(* IEC 61131-3 sources: rusty/tests/lit/single/type_promotion/bit_string/case_selector, 5 files *)

(* ---- byte_range_across_midpoint.st ---- *)
// RUN: %COMPILE %s && %RUN | %CHECK %s
// A range label that crosses the signed midpoint of the BYTE selector matches every value between its bounds.
FUNCTION branch : DINT
    VAR_INPUT
        x : BYTE;
    END_VAR

    CASE x OF
        16#00:
            branch := 1;
        16#01..16#09:
            branch := 2;
        16#0B..16#FE:
            branch := 3;
        16#FF:
            branch := 4;
    ELSE
        branch := 9;
    END_CASE
END_FUNCTION

FUNCTION main : DINT
    printf('16#00 -> %d$N', branch(16#00));                     // CHECK: 16#00 -> 1
    printf('16#05 -> %d$N', branch(16#05));                     // CHECK-NEXT: 16#05 -> 2
    printf('16#0A -> %d$N', branch(16#0A));                     // CHECK-NEXT: 16#0A -> 9
    printf('16#0B -> %d$N', branch(16#0B));                     // CHECK-NEXT: 16#0B -> 3
    printf('16#7F -> %d$N', branch(16#7F));                     // CHECK-NEXT: 16#7F -> 3
    printf('16#80 -> %d$N', branch(16#80));                     // CHECK-NEXT: 16#80 -> 3
    printf('16#C8 -> %d$N', branch(16#C8));                     // CHECK-NEXT: 16#C8 -> 3
    printf('16#FE -> %d$N', branch(16#FE));                     // CHECK-NEXT: 16#FE -> 3
    printf('16#FF -> %d$N', branch(16#FF));                     // CHECK-NEXT: 16#FF -> 4
END_FUNCTION

(* ---- dword_range_across_midpoint.st ---- *)
// RUN: %COMPILE %s && %RUN | %CHECK %s
// A range label that crosses the signed midpoint of the DWORD selector matches every value between its bounds.
FUNCTION branch : DINT
    VAR_INPUT
        x : DWORD;
    END_VAR

    CASE x OF
        16#0000_0000:
            branch := 1;
        16#0000_0001..16#0000_0009:
            branch := 2;
        16#0000_000B..16#FFFF_FFFE:
            branch := 3;
        16#FFFF_FFFF:
            branch := 4;
    ELSE
        branch := 9;
    END_CASE
END_FUNCTION

FUNCTION main : DINT
    printf('16#0000_0000 -> %d$N', branch(16#0000_0000));       // CHECK: 16#0000_0000 -> 1
    printf('16#0000_0005 -> %d$N', branch(16#0000_0005));       // CHECK-NEXT: 16#0000_0005 -> 2
    printf('16#0000_000A -> %d$N', branch(16#0000_000A));       // CHECK-NEXT: 16#0000_000A -> 9
    printf('16#0000_000B -> %d$N', branch(16#0000_000B));       // CHECK-NEXT: 16#0000_000B -> 3
    printf('16#7FFF_FFFF -> %d$N', branch(16#7FFF_FFFF));       // CHECK-NEXT: 16#7FFF_FFFF -> 3
    printf('16#8000_0000 -> %d$N', branch(16#8000_0000));       // CHECK-NEXT: 16#8000_0000 -> 3
    printf('16#B2D0_5E00 -> %d$N', branch(16#B2D0_5E00));       // CHECK-NEXT: 16#B2D0_5E00 -> 3
    printf('16#FFFF_FFFE -> %d$N', branch(16#FFFF_FFFE));       // CHECK-NEXT: 16#FFFF_FFFE -> 3
    printf('16#FFFF_FFFF -> %d$N', branch(16#FFFF_FFFF));       // CHECK-NEXT: 16#FFFF_FFFF -> 4
END_FUNCTION

(* ---- lword_range_across_midpoint.st ---- *)
// RUN: %COMPILE %s && %RUN | %CHECK %s
// A range label that crosses the signed midpoint of the LWORD selector matches every value between its bounds.
FUNCTION branch : DINT
    VAR_INPUT
        x : LWORD;
    END_VAR

    CASE x OF
        16#0:
            branch := 1;
        16#1..16#9:
            branch := 2;
        16#B..16#FFFF_FFFF_FFFF_FFFE:
            branch := 3;
        16#FFFF_FFFF_FFFF_FFFF:
            branch := 4;
    ELSE
        branch := 9;
    END_CASE
END_FUNCTION

FUNCTION main : DINT
    printf('16#0 -> %d$N', branch(16#0));                       // CHECK: 16#0 -> 1
    printf('16#5 -> %d$N', branch(16#5));                       // CHECK-NEXT: 16#5 -> 2
    printf('16#A -> %d$N', branch(16#A));                       // CHECK-NEXT: 16#A -> 9
    printf('16#B -> %d$N', branch(16#B));                       // CHECK-NEXT: 16#B -> 3
    printf('16#7FFF_FFFF_FFFF_FFFF -> %d$N', branch(16#7FFF_FFFF_FFFF_FFFF));  // CHECK-NEXT: 16#7FFF_FFFF_FFFF_FFFF -> 3
    printf('16#8000_0000_0000_0000 -> %d$N', branch(16#8000_0000_0000_0000));  // CHECK-NEXT: 16#8000_0000_0000_0000 -> 3
    printf('16#A000_0000_0000_0000 -> %d$N', branch(16#A000_0000_0000_0000));  // CHECK-NEXT: 16#A000_0000_0000_0000 -> 3
    printf('16#FFFF_FFFF_FFFF_FFFE -> %d$N', branch(16#FFFF_FFFF_FFFF_FFFE));  // CHECK-NEXT: 16#FFFF_FFFF_FFFF_FFFE -> 3
    printf('16#FFFF_FFFF_FFFF_FFFF -> %d$N', branch(16#FFFF_FFFF_FFFF_FFFF));  // CHECK-NEXT: 16#FFFF_FFFF_FFFF_FFFF -> 4
END_FUNCTION

(* ---- range_within_one_half.st ---- *)
// RUN: %COMPILE %s && %RUN | %CHECK %s
// Range labels that stay below or above the signed midpoint of a bit string selector.
FUNCTION branch_byte : DINT
    VAR_INPUT
        x : BYTE;
    END_VAR

    CASE x OF
        16#01..16#64: branch_byte := 1;
        16#81..16#FE: branch_byte := 2;
        16#FF: branch_byte := 3;
    ELSE
        branch_byte := 9;
    END_CASE
END_FUNCTION

FUNCTION branch_dword : DINT
    VAR_INPUT
        x : DWORD;
    END_VAR

    CASE x OF
        16#0000_0001..16#0000_FFFF: branch_dword := 1;
        16#8000_0000..16#FFFF_FFFE: branch_dword := 2;
        16#FFFF_FFFF: branch_dword := 3;
    ELSE
        branch_dword := 9;
    END_CASE
END_FUNCTION

FUNCTION main : DINT
    // BYTE
    printf('BYTE 16#32 -> %d$N', branch_byte(16#32));                   // CHECK: BYTE 16#32 -> 1
    printf('BYTE 16#C8 -> %d$N', branch_byte(16#C8));                   // CHECK-NEXT: BYTE 16#C8 -> 2
    printf('BYTE 16#FF -> %d$N', branch_byte(16#FF));                   // CHECK-NEXT: BYTE 16#FF -> 3

    // DWORD
    printf('DWORD 16#10 -> %d$N', branch_dword(16#10));                 // CHECK-NEXT: DWORD 16#10 -> 1
    printf('DWORD 16#8000_0001 -> %d$N', branch_dword(16#8000_0001));   // CHECK-NEXT: DWORD 16#8000_0001 -> 2
    printf('DWORD 16#FFFF_FFFF -> %d$N', branch_dword(16#FFFF_FFFF));   // CHECK-NEXT: DWORD 16#FFFF_FFFF -> 3
END_FUNCTION

(* ---- word_range_across_midpoint.st ---- *)
// RUN: %COMPILE %s && %RUN | %CHECK %s
// A range label that crosses the signed midpoint of the WORD selector matches every value between its bounds.
FUNCTION branch : DINT
    VAR_INPUT
        x : WORD;
    END_VAR

    CASE x OF
        16#0000:
            branch := 1;
        16#0001..16#0009:
            branch := 2;
        16#000B..16#FFFE:
            branch := 3;
        16#FFFF:
            branch := 4;
    ELSE
        branch := 9;
    END_CASE
END_FUNCTION

FUNCTION main : DINT
    printf('16#0000 -> %d$N', branch(16#0000));                 // CHECK: 16#0000 -> 1
    printf('16#0005 -> %d$N', branch(16#0005));                 // CHECK-NEXT: 16#0005 -> 2
    printf('16#000A -> %d$N', branch(16#000A));                 // CHECK-NEXT: 16#000A -> 9
    printf('16#000B -> %d$N', branch(16#000B));                 // CHECK-NEXT: 16#000B -> 3
    printf('16#7FFF -> %d$N', branch(16#7FFF));                 // CHECK-NEXT: 16#7FFF -> 3
    printf('16#8000 -> %d$N', branch(16#8000));                 // CHECK-NEXT: 16#8000 -> 3
    printf('16#9C40 -> %d$N', branch(16#9C40));                 // CHECK-NEXT: 16#9C40 -> 3
    printf('16#FFFE -> %d$N', branch(16#FFFE));                 // CHECK-NEXT: 16#FFFE -> 3
    printf('16#FFFF -> %d$N', branch(16#FFFF));                 // CHECK-NEXT: 16#FFFF -> 4
END_FUNCTION
